    PROC Path_RobotLab(PERS wobjdata WO_Pastel)
        Path_vacio_ejecucion p_vacio_labSIR, 1, WO_Pastel, FALSE;
        index_vacio_destino:=25;
        Path_contacto_ejecucion p_contacto_labSIR, 1, 3, WO_Pastel, FALSE;
        Mover_en_contacto;
        TriggC p_contacto_labSIR{4},p_contacto_labSIR{5},Vel_Proceso,triggContactoCir,Z_Proceso,Prototipo_JSDaleman\WObj:=WO_Pastel;
        TriggL p_contacto_labSIR{6},Vel_Proceso,triggContacto,Z_Proceso,Prototipo_JSDaleman\WObj:=WO_Pastel;
        TriggC p_contacto_labSIR{7},p_contacto_labSIR{8},Vel_Proceso,triggContactoCir,Z_Proceso,Prototipo_JSDaleman\WObj:=WO_Pastel;
        Path_contacto_ejecucion p_contacto_labSIR, 9, 25, WO_Pastel, TRUE;
        Path_vacio_ejecucion p_vacio_labSIR, 2, WO_Pastel, FALSE;
        Path_contacto_ejecucion p_contacto_labSIR, 26, 94, WO_Pastel, TRUE;
        Path_vacio_ejecucion p_vacio_labSIR, 3, WO_Pastel, FALSE;
        Path_contacto_ejecucion p_contacto_labSIR, 95, 111, WO_Pastel, TRUE;
        Path_vacio_ejecucion p_vacio_labSIR, 4, WO_Pastel, FALSE;
        Path_contacto_ejecucion p_contacto_labSIR, 112, 125, WO_Pastel, TRUE;
        Path_vacio_ejecucion p_vacio_labSIR, 5, WO_Pastel, FALSE;
        index_vacio_destino:=131;
        Mover_a_contacto;
        TriggL p_contacto_labSIR{126},Vel_Acercamiento,triggContacto,Z_Acercamiento,Prototipo_JSDaleman\WObj:=WO_Pastel;
        Mover_en_contacto;
        TriggC p_contacto_labSIR{127},p_contacto_labSIR{128},Vel_Proceso,triggContactoCir,Z_Proceso,Prototipo_JSDaleman\WObj:=WO_Pastel;
        TriggC p_contacto_labSIR{129},p_contacto_labSIR{130},Vel_Proceso,triggContactoCir,Z_Proceso,Prototipo_JSDaleman\WObj:=WO_Pastel;
        Mover_a_vacio;
        TriggL p_contacto_labSIR{131},Vel_Acercamiento,triggContacto,Z_Acercamiento,Prototipo_JSDaleman\WObj:=WO_Pastel;
        Path_vacio_ejecucion p_vacio_labSIR, 6, WO_Pastel, FALSE;
        index_vacio_destino:=137;
        Mover_a_contacto;
        TriggL p_contacto_labSIR{132},Vel_Acercamiento,triggContacto,Z_Acercamiento,Prototipo_JSDaleman\WObj:=WO_Pastel;
        Mover_en_contacto;
        TriggC p_contacto_labSIR{133},p_contacto_labSIR{134},Vel_Proceso,triggContactoCir,Z_Proceso,Prototipo_JSDaleman\WObj:=WO_Pastel;
        TriggC p_contacto_labSIR{135},p_contacto_labSIR{136},Vel_Proceso,triggContactoCir,Z_Proceso,Prototipo_JSDaleman\WObj:=WO_Pastel;
        Mover_a_vacio;
        TriggL p_contacto_labSIR{137},Vel_Acercamiento,triggContacto,Z_Acercamiento,Prototipo_JSDaleman\WObj:=WO_Pastel;
        Path_vacio_ejecucion p_vacio_labSIR, 7, WO_Pastel, FALSE;
        index_vacio_destino:=143;
        Mover_a_contacto;
        TriggL p_contacto_labSIR{138},Vel_Acercamiento,triggContacto,Z_Acercamiento,Prototipo_JSDaleman\WObj:=WO_Pastel;
        Mover_en_contacto;
        TriggC p_contacto_labSIR{139},p_contacto_labSIR{140},Vel_Proceso,triggContactoCir,Z_Proceso,Prototipo_JSDaleman\WObj:=WO_Pastel;
        TriggC p_contacto_labSIR{141},p_contacto_labSIR{142},Vel_Proceso,triggContactoCir,Z_Proceso,Prototipo_JSDaleman\WObj:=WO_Pastel;
        Mover_a_vacio;
        TriggL p_contacto_labSIR{143},Vel_Acercamiento,triggContacto,Z_Acercamiento,Prototipo_JSDaleman\WObj:=WO_Pastel;
        Path_vacio_ejecucion p_vacio_labSIR, 8, WO_Pastel, FALSE;
        index_vacio_destino:=149;
        Mover_a_contacto;
        TriggL p_contacto_labSIR{144},Vel_Acercamiento,triggContacto,Z_Acercamiento,Prototipo_JSDaleman\WObj:=WO_Pastel;
        Mover_en_contacto;
        TriggC p_contacto_labSIR{145},p_contacto_labSIR{146},Vel_Proceso,triggContactoCir,Z_Proceso,Prototipo_JSDaleman\WObj:=WO_Pastel;
        TriggC p_contacto_labSIR{147},p_contacto_labSIR{148},Vel_Proceso,triggContactoCir,Z_Proceso,Prototipo_JSDaleman\WObj:=WO_Pastel;
        Mover_a_vacio;
        TriggL p_contacto_labSIR{149},Vel_Acercamiento,triggContacto,Z_Acercamiento,Prototipo_JSDaleman\WObj:=WO_Pastel;
        Path_vacio_ejecucion p_vacio_labSIR, 9, WO_Pastel, FALSE;
        index_vacio_destino:=155;
        Mover_a_contacto;
        TriggL p_contacto_labSIR{150},Vel_Acercamiento,triggContacto,Z_Acercamiento,Prototipo_JSDaleman\WObj:=WO_Pastel;
        Mover_en_contacto;
        TriggC p_contacto_labSIR{151},p_contacto_labSIR{152},Vel_Proceso,triggContactoCir,Z_Proceso,Prototipo_JSDaleman\WObj:=WO_Pastel;
        TriggC p_contacto_labSIR{153},p_contacto_labSIR{154},Vel_Proceso,triggContactoCir,Z_Proceso,Prototipo_JSDaleman\WObj:=WO_Pastel;
        Mover_a_vacio;
        TriggL p_contacto_labSIR{155},Vel_Acercamiento,triggContacto,Z_Acercamiento,Prototipo_JSDaleman\WObj:=WO_Pastel;
        Path_vacio_ejecucion p_vacio_labSIR, 10, WO_Pastel, FALSE;
        index_vacio_destino:=161;
        Mover_a_contacto;
        TriggL p_contacto_labSIR{156},Vel_Acercamiento,triggContacto,Z_Acercamiento,Prototipo_JSDaleman\WObj:=WO_Pastel;
        Mover_en_contacto;
        TriggC p_contacto_labSIR{157},p_contacto_labSIR{158},Vel_Proceso,triggContactoCir,Z_Proceso,Prototipo_JSDaleman\WObj:=WO_Pastel;
        TriggC p_contacto_labSIR{159},p_contacto_labSIR{160},Vel_Proceso,triggContactoCir,Z_Proceso,Prototipo_JSDaleman\WObj:=WO_Pastel;
        Mover_a_vacio;
        TriggL p_contacto_labSIR{161},Vel_Proceso,triggContacto,Z_Proceso,Prototipo_JSDaleman\WObj:=WO_Pastel;
    ENDPROC
    PROC Path_Tapa_LabSIR(PERS wobjdata WO_Pastel)
        Mover_en_vacio;
        MoveJ Target_Home_10,Vel_Vacio_Rap,Z_Vacio_Rap,Prototipo_JSDaleman\WObj:=wobj0;
        ReiniciarIndices;
        path_contacto_actual:="p_contacto_labSIR";
        path_vacio_actual:="p_vacio_labSIR";
        Path_RobotLab WO_Pastel;
        Path_LabSIR WO_Pastel;
        Mover_en_vacio;
        MoveJ Target_Home_10,Vel_Vacio_Rap,Z_Vacio_Rap,Prototipo_JSDaleman\WObj:=wobj0;
    ENDPROC
    PROC Path_LabSIR(PERS wobjdata WO_Pastel)
        Path_vacio_ejecucion p_vacio_labSIR, 11, WO_Pastel, FALSE;
        Path_contacto_ejecucion p_contacto_labSIR, 162, 170, WO_Pastel, TRUE;
        Path_vacio_ejecucion p_vacio_labSIR, 12, WO_Pastel, FALSE;
        Path_contacto_ejecucion p_contacto_labSIR, 171, 182, WO_Pastel, TRUE;
        Path_vacio_ejecucion p_vacio_labSIR, 13, WO_Pastel, FALSE;
        Path_contacto_ejecucion p_contacto_labSIR, 183, 188, WO_Pastel, TRUE;
        Path_vacio_ejecucion p_vacio_labSIR, 14, WO_Pastel, FALSE;
        Path_contacto_ejecucion p_contacto_labSIR, 189, 199, WO_Pastel, TRUE;
        Path_vacio_ejecucion p_vacio_labSIR, 15, WO_Pastel, FALSE;
        Path_contacto_ejecucion p_contacto_labSIR, 200, 205, WO_Pastel, TRUE;
        Path_vacio_ejecucion p_vacio_labSIR, 16, WO_Pastel, FALSE;
        Path_contacto_ejecucion p_contacto_labSIR, 206, 219, WO_Pastel, TRUE;
        Path_vacio_ejecucion p_vacio_labSIR, 17, WO_Pastel, FALSE;
        Path_contacto_ejecucion p_contacto_labSIR, 220, 226, WO_Pastel, TRUE;
        Path_vacio_ejecucion p_vacio_labSIR, 18, WO_Pastel, FALSE;
        Path_contacto_ejecucion p_contacto_labSIR, 227, 232, WO_Pastel, TRUE;
        Path_vacio_ejecucion p_vacio_labSIR, 19, WO_Pastel, FALSE;
        Path_contacto_ejecucion p_contacto_labSIR, 233, 256, WO_Pastel, TRUE;
    ENDPROC
    PROC Path_Frente_LabSIR(PERS wobjdata WO_Pastel)
        Mover_en_vacio;
        MoveJ Target_Home_10,Vel_Vacio_Rap,Z_Vacio_Rap,Prototipo_JSDaleman\WObj:=wobj0;
        MoveJ Target_Frente_10,Vel_Vacio,Z_VacioMov,Prototipo_JSDaleman\WObj:=WO_Pastel;
        MoveJ Target_Frente_20,Vel_Vacio,Z_VacioMov,Prototipo_JSDaleman\WObj:=WO_Pastel;
        ReiniciarIndices;
        path_contacto_actual:="p_contacto_labSIR_FrenteL";
        path_vacio_actual:="p_vacio_labSIR_FrenteL";
        Path_Chip WO_Pastel;
        Path_LetreroFrontal1_LabSIR WO_Pastel;
        Path_LetreroFrontal2_LabSIR WO_Pastel;
        Mover_en_vacio;
        MoveJ Target_Frente_20,Vel_Vacio,Z_VacioMov,Prototipo_JSDaleman\WObj:=WO_Pastel;
        MoveJ Target_Frente_10,Vel_Vacio,Z_VacioMov,Prototipo_JSDaleman\WObj:=WO_Pastel;
        MoveJ Target_Home_10,Vel_Vacio_Rap,Z_Vacio_Rap,Prototipo_JSDaleman\WObj:=wobj0;
        MoveJ Target_Frente_30,Vel_Vacio_Rap,Z_Vacio_Rap,Prototipo_JSDaleman\WObj:=WO_Pastel;
        MoveJ Target_Frente_40,Vel_Vacio_Rap,Z_Vacio_Rap,Prototipo_JSDaleman\WObj:=WO_Pastel;
        ReiniciarIndices;
        path_contacto_actual:="p_contacto_labSIR_FrenteR";
        path_vacio_actual:="p_vacio_labSIR_FrenteR";
        Path_Engranaje WO_Pastel;
        Path_LetreroFrontal3_LabSIR WO_Pastel;
        Path_LetreroFrontal4_LabSIR WO_Pastel;
        Mover_en_vacio;
        MoveJ Target_Frente_40,Vel_Vacio_Rap,Z_Vacio_Rap,Prototipo_JSDaleman\WObj:=WO_Pastel;
        MoveJ Target_Frente_30,Vel_Vacio_Rap,Z_Vacio_Rap,Prototipo_JSDaleman\WObj:=WO_Pastel;
        MoveJ Target_Home_10,Vel_Vacio_Rap,Z_Vacio_Rap,Prototipo_JSDaleman\WObj:=wobj0;
    ENDPROC
    PROC Path_Chip(PERS wobjdata WO_Pastel)
        Path_vacio_ejecucion p_vacio_labSIR_FrenteL, 1, WO_Pastel, FALSE;
        Path_contacto_ejecucion p_contacto_labSIR_FrenteL, 1, 50, WO_Pastel, TRUE;
        Path_vacio_ejecucion p_vacio_labSIR_FrenteL, 1, WO_Pastel, FALSE;
        Path_contacto_ejecucion p_contacto_labSIR_FrenteL, 51, 56, WO_Pastel, TRUE;
    ENDPROC
    PROC Path_LetreroFrontal1_LabSIR(PERS wobjdata WO_Pastel)
        Path_vacio_ejecucion p_vacio_labSIR_FrenteL, 3, WO_Pastel, FALSE;
        Path_contacto_ejecucion p_contacto_labSIR_FrenteL, 57, 60, WO_Pastel, TRUE;
        Path_vacio_ejecucion p_vacio_labSIR_FrenteL, 4, WO_Pastel, FALSE;
        Path_contacto_ejecucion p_contacto_labSIR_FrenteL, 61, 74, WO_Pastel, TRUE;
        Path_vacio_ejecucion p_vacio_labSIR_FrenteL, 5, WO_Pastel, FALSE;
        Path_contacto_ejecucion p_contacto_labSIR_FrenteL, 75, 92, WO_Pastel, TRUE;
        Path_vacio_ejecucion p_vacio_labSIR_FrenteL, 6, WO_Pastel, FALSE;
        Path_contacto_ejecucion p_contacto_labSIR_FrenteL, 93, 116, WO_Pastel, TRUE;
        Path_vacio_ejecucion p_vacio_labSIR_FrenteL, 7, WO_Pastel, FALSE;
        Path_contacto_ejecucion p_contacto_labSIR_FrenteL, 117, 122, WO_Pastel, TRUE;
        Path_vacio_ejecucion p_vacio_labSIR_FrenteL, 8, WO_Pastel, FALSE;
        Path_contacto_ejecucion p_contacto_labSIR_FrenteL, 123, 140, WO_Pastel, TRUE;
        Path_vacio_ejecucion p_vacio_labSIR_FrenteL, 9, WO_Pastel, FALSE;
        Path_contacto_ejecucion p_contacto_labSIR_FrenteL, 141, 149, WO_Pastel, TRUE;
        Path_vacio_ejecucion p_vacio_labSIR_FrenteL, 10, WO_Pastel, FALSE;
        Path_contacto_ejecucion p_contacto_labSIR_FrenteL, 150, 174, WO_Pastel, TRUE;
        Path_vacio_ejecucion p_vacio_labSIR_FrenteL, 11, WO_Pastel, FALSE;
        Path_contacto_ejecucion p_contacto_labSIR_FrenteL, 175, 183, WO_Pastel, TRUE;
        Path_vacio_ejecucion p_vacio_labSIR_FrenteL, 12, WO_Pastel, FALSE;
        Path_contacto_ejecucion p_contacto_labSIR_FrenteL, 184, 186, WO_Pastel, TRUE;
        Path_vacio_ejecucion p_vacio_labSIR_FrenteL, 13, WO_Pastel, FALSE;
        index_vacio_destino:=188;
        Mover_a_contacto;
        TriggL p_contacto_labSIR_FrenteL{187},Vel_Acercamiento,triggContacto,Z_Acercamiento,Prototipo_JSDaleman\WObj:=WO_Pastel;
        Mover_en_contacto;
        TriggL p_contacto_labSIR_FrenteL{188},Vel_Acercamiento_Lateral,triggContacto,Z_Acercamiento,Prototipo_JSDaleman\WObj:=WO_Pastel;
        Path_vacio_ejecucion p_vacio_labSIR_FrenteL, 14, WO_Pastel, FALSE;
        Path_contacto_ejecucion p_contacto_labSIR_FrenteL, 189, 212, WO_Pastel, TRUE;
    ENDPROC
    PROC Path_LetreroFrontal2_LabSIR(PERS wobjdata WO_Pastel)
        Path_vacio_ejecucion p_vacio_labSIR_FrenteL, 15, WO_Pastel, FALSE;
        Path_contacto_ejecucion p_contacto_labSIR_FrenteL, 213, 238, WO_Pastel, TRUE;
        Path_vacio_ejecucion p_vacio_labSIR_FrenteL, 16, WO_Pastel, FALSE;
        Path_contacto_ejecucion p_contacto_labSIR_FrenteL, 239, 262, WO_Pastel, TRUE;
        Path_vacio_ejecucion p_vacio_labSIR_FrenteL, 17, WO_Pastel, FALSE;
        Path_contacto_ejecucion p_contacto_labSIR_FrenteL, 263, 273, WO_Pastel, TRUE;
        Path_vacio_ejecucion p_vacio_labSIR_FrenteL, 18, WO_Pastel, FALSE;
        Path_contacto_ejecucion p_contacto_labSIR_FrenteL, 274, 287, WO_Pastel, TRUE;
        Path_vacio_ejecucion p_vacio_labSIR_FrenteL, 19, WO_Pastel, FALSE;
        Path_contacto_ejecucion p_contacto_labSIR_FrenteL, 288, 307, WO_Pastel, TRUE;
        Path_vacio_ejecucion p_vacio_labSIR_FrenteL, 20, WO_Pastel, FALSE;
        Path_contacto_ejecucion p_contacto_labSIR_FrenteL, 308, 341, WO_Pastel, TRUE;
        Path_vacio_ejecucion p_vacio_labSIR_FrenteL, 21, WO_Pastel, FALSE;
        Path_contacto_ejecucion p_contacto_labSIR_FrenteL, 342, 344, WO_Pastel, TRUE;
        Path_vacio_ejecucion p_vacio_labSIR_FrenteL, 22, WO_Pastel, FALSE;
        Path_contacto_ejecucion p_contacto_labSIR_FrenteL, 345, 346, WO_Pastel, TRUE;
        Path_vacio_ejecucion p_vacio_labSIR_FrenteL, 23, WO_Pastel, FALSE;
        Path_contacto_ejecucion p_contacto_labSIR_FrenteL, 347, 350, WO_Pastel, TRUE;
        Path_vacio_ejecucion p_vacio_labSIR_FrenteL, 24, WO_Pastel, FALSE;
        Path_contacto_ejecucion p_contacto_labSIR_FrenteL, 351, 370, WO_Pastel, TRUE;
        Path_vacio_ejecucion p_vacio_labSIR_FrenteL, 25, WO_Pastel, FALSE;
        Path_contacto_ejecucion p_contacto_labSIR_FrenteL, 371, 379, WO_Pastel, TRUE;
        Path_vacio_ejecucion p_vacio_labSIR_FrenteL, 26, WO_Pastel, FALSE;
        Path_contacto_ejecucion p_contacto_labSIR_FrenteL, 380, 391, WO_Pastel, TRUE;
        Path_vacio_ejecucion p_vacio_labSIR_FrenteL, 27, WO_Pastel, FALSE;
        Path_contacto_ejecucion p_contacto_labSIR_FrenteL, 392, 394, WO_Pastel, TRUE;
    ENDPROC
    PROC Path_Engranaje(PERS wobjdata WO_Pastel)
        Path_vacio_ejecucion p_vacio_labSIR_FrenteR, 1, WO_Pastel, FALSE;
        Path_contacto_ejecucion p_contacto_labSIR_FrenteR, 1, 78, WO_Pastel, TRUE;
        Path_vacio_ejecucion p_vacio_labSIR_FrenteR, 2, WO_Pastel, FALSE;
        Path_contacto_ejecucion p_contacto_labSIR_FrenteR, 79, 97, WO_Pastel, TRUE;
    ENDPROC
    PROC Path_LetreroFrontal3_LabSIR(PERS wobjdata WO_Pastel)
        Path_vacio_ejecucion p_vacio_labSIR_FrenteR, 3, WO_Pastel, FALSE;
        Path_contacto_ejecucion p_contacto_labSIR_FrenteR, 98, 121, WO_Pastel, TRUE;
        Path_vacio_ejecucion p_vacio_labSIR_FrenteR, 4, WO_Pastel, FALSE;
        Path_contacto_ejecucion p_contacto_labSIR_FrenteR, 122, 150, WO_Pastel, TRUE;
        Path_vacio_ejecucion p_vacio_labSIR_FrenteR, 5, WO_Pastel, FALSE;
        Path_contacto_ejecucion p_contacto_labSIR_FrenteR, 151, 163, WO_Pastel, TRUE;
        Path_vacio_ejecucion p_vacio_labSIR_FrenteR, 6, WO_Pastel, FALSE;
        Path_contacto_ejecucion p_contacto_labSIR_FrenteR, 164, 187, WO_Pastel, TRUE;
        Path_vacio_ejecucion p_vacio_labSIR_FrenteR, 7, WO_Pastel, FALSE;
        Path_contacto_ejecucion p_contacto_labSIR_FrenteR, 188, 198, WO_Pastel, TRUE;
        Path_vacio_ejecucion p_vacio_labSIR_FrenteR, 8, WO_Pastel, FALSE;
        Path_contacto_ejecucion p_contacto_labSIR_FrenteR, 199, 218, WO_Pastel, TRUE;
        Path_vacio_ejecucion p_vacio_labSIR_FrenteR, 9, WO_Pastel, FALSE;
        Path_contacto_ejecucion p_contacto_labSIR_FrenteR, 219, 221, WO_Pastel, TRUE;
        Path_vacio_ejecucion p_vacio_labSIR_FrenteR, 10, WO_Pastel, FALSE;
        Path_contacto_ejecucion p_contacto_labSIR_FrenteR, 222, 223, WO_Pastel, TRUE;
        Path_vacio_ejecucion p_vacio_labSIR_FrenteR, 11, WO_Pastel, FALSE;
        Path_contacto_ejecucion p_contacto_labSIR_FrenteR, 224, 242, WO_Pastel, TRUE;
        Path_vacio_ejecucion p_vacio_labSIR_FrenteR, 12, WO_Pastel, FALSE;
        Path_contacto_ejecucion p_contacto_labSIR_FrenteR, 243, 264, WO_Pastel, TRUE;
        Path_vacio_ejecucion p_vacio_labSIR_FrenteR, 13, WO_Pastel, FALSE;
        Path_contacto_ejecucion p_contacto_labSIR_FrenteR, 265, 281, WO_Pastel, TRUE;
    ENDPROC
    PROC Path_LetreroFrontal4_LabSIR(PERS wobjdata WO_Pastel)
        Path_vacio_ejecucion p_vacio_labSIR_FrenteR, 14, WO_Pastel, FALSE;
        Path_contacto_ejecucion p_contacto_labSIR_FrenteR, 282, 293, WO_Pastel, TRUE;
        Path_vacio_ejecucion p_vacio_labSIR_FrenteR, 15, WO_Pastel, FALSE;
        Path_contacto_ejecucion p_contacto_labSIR_FrenteR, 294, 317, WO_Pastel, TRUE;
        Path_vacio_ejecucion p_vacio_labSIR_FrenteR, 16, WO_Pastel, FALSE;
        Path_contacto_ejecucion p_contacto_labSIR_FrenteR, 318, 332, WO_Pastel, TRUE;
        Path_vacio_ejecucion p_vacio_labSIR_FrenteR, 17, WO_Pastel, FALSE;
        Path_contacto_ejecucion p_contacto_labSIR_FrenteR, 333, 350, WO_Pastel, TRUE;
        Path_vacio_ejecucion p_vacio_labSIR_FrenteR, 18, WO_Pastel, FALSE;
        Path_contacto_ejecucion p_contacto_labSIR_FrenteR, 351, 360, WO_Pastel, TRUE;
        Path_vacio_ejecucion p_vacio_labSIR_FrenteR, 19, WO_Pastel, FALSE;
        Path_contacto_ejecucion p_contacto_labSIR_FrenteR, 361, 363, WO_Pastel, TRUE;
        Path_vacio_ejecucion p_vacio_labSIR_FrenteR, 20, WO_Pastel, FALSE;
        Path_contacto_ejecucion p_contacto_labSIR_FrenteR, 364, 365, WO_Pastel, TRUE;
        Path_vacio_ejecucion p_vacio_labSIR_FrenteR, 21, WO_Pastel, FALSE;
        Path_contacto_ejecucion p_contacto_labSIR_FrenteR, 366, 370, WO_Pastel, TRUE;
        Path_vacio_ejecucion p_vacio_labSIR_FrenteR, 22, WO_Pastel, FALSE;
        Path_contacto_ejecucion p_contacto_labSIR_FrenteR, 371, 394, WO_Pastel, TRUE;
        Path_vacio_ejecucion p_vacio_labSIR_FrenteR, 23, WO_Pastel, FALSE;
        Path_contacto_ejecucion p_contacto_labSIR_FrenteR, 395, 410, WO_Pastel, TRUE;
        Path_vacio_ejecucion p_vacio_labSIR_FrenteR, 24, WO_Pastel, FALSE;
        Path_contacto_ejecucion p_contacto_labSIR_FrenteR, 411, 430, WO_Pastel, TRUE;
        Path_vacio_ejecucion p_vacio_labSIR_FrenteR, 25, WO_Pastel, FALSE;
        Path_contacto_ejecucion p_contacto_labSIR_FrenteR, 431, 448, WO_Pastel, TRUE;
    ENDPROC
ENDMODULE
